(* IEC 61131-3 sources: volt/packages/volt-lsp-iec/test-corpus/pro2193/Device/Plc Logic/Application/09 Misc/Library Manager/L_TB1P_TechnologyBasics, 21 files *)

(* ---- L_TB1P_DIRECTION.dut ---- *)
TYPE L_TB1P_DIRECTION :
(
	DEFAULT := 0,
	CW := 1,
	CCW := 2
);
END_TYPE

(* ---- L_TB1P_STATES.dut ---- *)
TYPE L_TB1P_STATES :
(
	INIT := 1,
	READY := 2,
	CAMMING := 112,
	CAMMING_DONE := 113,
	CLUTCH_OPEN_INSTANT := 114,
	CLUTCH_CLOSE := 115,
	CLUTCH_OPEN := 116,
	CAMSEQUENCER_LOADCAMTABLE := 150,
	CAMSEQUENCER_CYCLICCAM1 := 151,
	CAMSEQUENCER_CYCLICCAM3 := 152,
	CAMSEQUENCER_CAM1CYCLICCAM3CAM1 := 153,
	CAMSEQUENCER_CAM1CAM2CYCLICCAM3CAM4CAM1 := 154,
	ERROR := 999
);
END_TYPE

(* ---- L_TB1P_CONSTANTS.gvl ---- *)
VAR_GLOBAL
	GC_POSITIVE_LIMIT_32BIT : LREAL := 2147483647;
	GC_NEGATIVE_LIMIT_32BIT : LREAL := -2147483647;
END_VAR

(* ---- GETBOOLEANPROPERTY.pou ---- *)
FUNCTION GETBOOLEANPROPERTY : BOOL
VAR_INPUT
	STKEY : WSTRING;
END_VAR
END_FUNCTION

(* ---- GETCOMPANY.pou ---- *)
FUNCTION GETCOMPANY : WSTRING
END_FUNCTION

(* ---- GETNUMBERPROPERTY.pou ---- *)
FUNCTION GETNUMBERPROPERTY : DINT
VAR_INPUT
	STKEY : WSTRING;
END_VAR
END_FUNCTION

(* ---- GETTEXTPROPERTY.pou ---- *)
FUNCTION GETTEXTPROPERTY : WSTRING
VAR_INPUT
	STKEY : WSTRING;
END_VAR
END_FUNCTION

(* ---- GETTEXTPROPERTY2.pou ---- *)
FUNCTION GETTEXTPROPERTY2 : POINTER TO WSTRING
VAR_INPUT
	STKEY : WSTRING;
END_VAR
END_FUNCTION

(* ---- GETTITLE.pou ---- *)
FUNCTION GETTITLE : WSTRING
END_FUNCTION

(* ---- GETVERSION.pou ---- *)
FUNCTION GETVERSION : VERSION
END_FUNCTION

(* ---- GETVERSIONPROPERTY.pou ---- *)
FUNCTION GETVERSIONPROPERTY : VERSION
VAR_INPUT
	STKEY : WSTRING;
END_VAR
END_FUNCTION

(* ---- GLOBALTEXTLIST.pou ---- *)
FUNCTION_BLOCK GLOBALTEXTLIST
VAR
	M_TEXTLISTFILE : STRING(255);
	_STNAMESPACE : STRING;
END_VAR
END_FUNCTION_BLOCK

(* ---- IMAGEPOOL.pou ---- *)
FUNCTION_BLOCK IMAGEPOOL
VAR
	M_STNAMESPACE : STRING(80);
	M_STHELPVARID : STRING;
	M_STHELPVARPATH : STRING(255);
	M_STHELP : STRING;
	M_REGISTERIMAGES : BOOL := TRUE;
END_VAR
END_FUNCTION_BLOCK

METHOD FB_INIT : BOOL
VAR_INPUT
	BINITRETAINS : BOOL;
	BINCOPYCODE : BOOL;
END_VAR
END_METHOD

METHOD FB_REINIT : BOOL
END_METHOD

METHOD FB_EXIT : BOOL
VAR_INPUT
	BINCOPYCODE : BOOL;
END_VAR
END_METHOD

(* ---- L_TB1P_ACCCOMP.pou ---- *)
FUNCTION_BLOCK L_TB1P_ACCCOMP
VAR_INPUT
	LRCYCVEL : LREAL;
	LRMINERTIAMAX : LREAL;
	LRMINERTIACONST : LREAL;
	LRVARIABLEMINERTIA : LREAL;
	LRMINERTIAADAPT : LREAL := 1.0;
	LRFILTERTIMEACCSPEED : REAL := 0.0;
	LRDEADBANDACCTORQUE : LREAL := 0.0;
	LRGAINPOS : LREAL := 1.0;
	LRGAINNEG : LREAL := 1.0;
	XRESET : BOOL;
END_VAR
VAR_OUTPUT
	LRSETACCOUT : LREAL;
	LRSETTORQUEOUT : LREAL;
END_VAR
VAR
	TBDIFFERENTIATE1 : L_USPP_Differentiate;
	LRMINERTIAVAR : LREAL;
	LRLRSETACC_INT : LREAL;
	LRFACTOR_INT : LREAL := 1;
	LRFACTOR : LREAL;
END_VAR
END_FUNCTION_BLOCK

(* ---- L_TB1P_CALCDIAMETER.pou ---- *)
FUNCTION_BLOCK L_TB1P_CALCDIAMETER
VAR_INPUT
	LRCYCREELSPEED : LREAL;
	LRCYCLINEVEL : LREAL;
	LRMAXDIAMETER : LREAL;
	LRMINDIAMETER : LREAL;
	LRCALCULATIONDISTANCE : LREAL := 1;
	XFORCECALCULATION : BOOL;
	XHOLDDIAMETER : BOOL;
	XUNIDIRECT : BOOL;
	XUNWINDACTIVE : BOOL;
	XLOADSETDIAMETER : BOOL;
	LRSETDIAMETER : LREAL;
	LRFILTERTIMEDIAMETER : LREAL := 0;
	LRWINDOWWEBBREAKMONIT : LREAL := 0.1;
END_VAR
VAR_OUTPUT
	XERROR : BOOL;
	EERRORID : L_IE1P_Error;
	LRSETDIAMETEROUT : LREAL;
	LRSETDIAMETERPCTOUT : LREAL;
	LRREZIPRDIAMETERPCT : LREAL;
	XDIAMETERMAXLIMIT : BOOL := FALSE;
	XDIAMETERMINLIMIT : BOOL := FALSE;
	XWEBBREAK : BOOL := FALSE;
	LRMINDIAMETERPCT : LREAL;
	LRSETMINERTIASCALEDOUT : LREAL;
END_VAR
VAR_IN_OUT
	LRDIAMETERRETAIN : LREAL := 0;
END_VAR
VAR
	LRTASKCYCLE : LREAL;
	XTASKCYCLEVALID : BOOL;
	LRFILTERTIME : LREAL;
	LRUNFILTEREDDIAMETER : LREAL;
	LRCALCULATIONDISTANCE_INT : LREAL;
	LRACTSPEEDREEL : LREAL;
	LRNWINDER : LREAL;
	LRREELPOSDIFF : LREAL;
	LRACTPOSDIFF : LREAL;
	LRACTLINESPEED : LREAL;
	LRWICKELWELLENDIFFERENZ : LREAL;
	LRCYCVELLINETMP : LREAL;
	LRSTOREDIAMETER : LREAL;
	LRDIAMETERMONITOR : LREAL;
	LRDIAMETERUNFILTERED : LREAL;
	LRTEMP : LREAL;
	LRTIME : LREAL;
	LRDMAXHYST : LREAL;
	LRDMINHYST : LREAL;
	XRESETCALCINTEGRATORFLAG : BOOL;
	LRMAXDIAMETERINT : LREAL;
	LRMAXDIAMETERMEM : LREAL;
	LRMINDIAMETERINT : LREAL;
	XRETAINLOCAL : BOOL := FALSE;
	LRDIAMETERINT : LREAL;
	LRREFDIAMWEBBREAK : LREAL;
	LRREFDIAMWEBBREAKSCALED : LREAL;
	LRCALCDISTLINEVEL_INT : LREAL;
	LRDIAMETER4CALCDIST : LREAL;
	LRCALCULATIONDISTANCE_OLD : LREAL;
	XHOLDINTEGRATOR_INT : BOOL;
	C_MINDIAMETER : LREAL := 1E-06;
	C_MAXDIAMETER : LREAL := 1000000.0;
	LRLINEVELINTEGRATED : LREAL;
	LRREFDIAMETERWEBBREAK : LREAL;
	LRSETDIAMETERUNFILTERED : LREAL;
	LRWINDERSPEEDINTEGRATED : LREAL;
	XDIAMCALCULATED : BOOL;
	XHOLDINTEGRATOR : BOOL;
END_VAR
END_FUNCTION_BLOCK

METHOD D_MIN_MAX
END_METHOD

METHOD LIMITER
END_METHOD

METHOD SETDIAMETER
VAR_INPUT
	LRNEWDIAMETER : LREAL;
END_VAR
END_METHOD

METHOD FB_INIT : BOOL
VAR_INPUT
	BINITRETAINS : BOOL;
	BINCOPYCODE : BOOL;
END_VAR
END_METHOD

(* ---- L_TB1P_FRICTIONCOMPENSATION.pou ---- *)
FUNCTION_BLOCK L_TB1P_FRICTIONCOMPENSATION
VAR_INPUT
	XIDENT : BOOL;
	XFOLLOWERACTIVE : BOOL;
	LRACTREELSPEEDIN : LREAL;
	LRACTTORQUEIN : LREAL;
	DWSELECTCURVE : DWORD;
	XENABLEFRICTIONCURVE : BOOL;
	LRSETREELSPEED : LREAL;
	LRFRICTIONADAPT : LREAL := 1;
	XINVERTOUTPUT : BOOL;
	LRMAXSPEEDIDENT : LREAL := 10;
	LRACCDECIDENT : LREAL := 1;
	LRFILTERTIMESPEED : LREAL := 0.005;
	LRFILTERTIMETORQUE : LREAL := 0.005;
	LRFILTERTIMEREELSPEED : LREAL := 0.0;
	LRLINEARCOMPSTART : LREAL;
	LRLINEARCOMPEND : LREAL;
	LRLINEARCOMPENDREELSPEED : LREAL;
END_VAR
VAR_OUTPUT
	XBUSY : BOOL;
	XDONE : BOOL;
	XERROR : BOOL := FALSE;
	EERRORID : L_IE1P_Error;
	XSTOP : BOOL;
	XENABLEFOLLOWER : BOOL;
	LRSETREELSPEEDOUT : LREAL;
	LRSETFRICTIONTORQUEOUT : LREAL;
END_VAR
VAR_IN_OUT
	ALRFRICTIONCURVE1 : ARRAY [1..66] OF LREAL;
	ALRFRICTIONCURVE2 : ARRAY [1..66] OF LREAL;
	ALRFRICTIONCURVE3 : ARRAY [1..66] OF LREAL;
	ALRFRICTIONCURVE4 : ARRAY [1..66] OF LREAL;
END_VAR
VAR
	LRTASKCYCLE : LREAL;
	DWINTERNALSTATE : DWORD;
	LRWINDOW : LREAL := 0.001;
	DISTATE : DINT;
	DWFRCURVENO : DWORD;
	XIMPOFF : BOOL;
	XFRICTIONBUSY : BOOL;
	XSTARTFRENABLE : BOOL;
	LRNACTFILTER : LREAL;
	LRMACTFILTER : LREAL;
	LRRAMPVALUE : LREAL;
	LRSTEP : LREAL;
	DWINDEX : DWORD;
	DWNUMBER : DWORD;
	ALRFRICTIONDATA1 : ARRAY [0..64] OF LREAL;
	ALRFRICTIONDATA2 : ARRAY [0..64] OF LREAL;
	LRDIST : LREAL;
	LRHALFDIST : LREAL;
	LRTEMP1 : LREAL;
	LRTEMP2 : LREAL;
	LRNMAXFRICTIONINT : LREAL;
	LRDIFFRAMP : LREAL;
	LRNMAXTIME : LREAL;
	LRACCDECIDENTINT : LREAL;
	LRTIME : LREAL;
	XENABLEFOLLOWEROLD : BOOL;
	LRSPEEDSETFILTER : LREAL;
	LRSPEEDSETFILTERABS : LREAL;
	LRSPEEDSETLIM : LREAL;
	LRDIFFFILTER : LREAL;
	LRACTFRICTION : LREAL;
	LRXTABLEVALUE : LREAL;
	LRMAXVALUE : LREAL;
	LRRESIDUAL : LREAL;
	LRSTRICH : LREAL;
	LRDELTAPOS : LREAL;
END_VAR
END_FUNCTION_BLOCK

METHOD RESETERROR
END_METHOD

(* ---- L_TB1P_IDENTMINERTIA.pou ---- *)
FUNCTION_BLOCK L_TB1P_IDENTMINERTIA
VAR_INPUT
	XIDENT : BOOL;
	XFOLLOWERACTIVE : BOOL;
	LRACTREELSPEEDIN : LREAL;
	LRACTTORQUEIN : LREAL;
	LRMAXSPEEDIDENT : LREAL := 10;
	LRMAXTORQUEIDENT : LREAL := 1;
	LRFILTERTIMESPEED : LREAL := 0.005;
	LRFILTERTIMETORQUE : LREAL := 0.005;
	LRFILTERTIMEREELSPEED : LREAL := 0.0;
END_VAR
VAR_OUTPUT
	XBUSY : BOOL;
	XDONE : BOOL;
	XERROR : BOOL := FALSE;
	EERRORID : L_IE1P_Error;
	XENABLEFOLLOWER : BOOL;
	LRSETTORQUEOUT : LREAL;
	LRMINERTIAIDENT : LREAL;
END_VAR
VAR
	LRMINERTIAMAXTOLERANCEERROR : LREAL;
	LRTASKCYCLE : LREAL;
	DWINTERNALSTATE : DWORD;
	DWINDEX : DWORD;
	DISTATE : DINT;
	XIMPOFF : BOOL;
	XACTIVE : BOOL;
	XMINERTIABUSY : BOOL;
	LRNACTFILTER : LREAL;
	LRMACTFILTER : LREAL;
	LRTIME : LREAL;
	LRNMAXMOTORINTERN : LREAL;
	LRMMAXMOTORINTERN : LREAL;
	LRNACTAKKU : LREAL;
	LRMACTAKKU : LREAL;
	LRSIGNNMAX : LREAL := 1;
	LRMSETMINERTIAINT_N : LREAL;
	LRNMAXMINERTIAINT_N : LREAL;
	LRACCTIME : LREAL;
	LRDECTIME : LREAL;
	LRTOTALTIME : LREAL;
	LRWAITTIME : LREAL;
END_VAR
END_FUNCTION_BLOCK

METHOD RESETERROR
END_METHOD

(* ---- L_TB1P_MARKREGISTER.pou ---- *)
FUNCTION_BLOCK L_TB1P_MARKREGISTER
VAR_INPUT
	XENABLE : BOOL;
	LRCYCSETVEL : LREAL;
	XTPRECEIVEDIN : BOOL;
	LRSETTPDIFFERENCE : LREAL;
	LRMARKSTACKLENGTH : LREAL;
	XCORRECTIONBUSY : BOOL;
	LRSETPOSCORRIN : LREAL;
END_VAR
VAR_OUTPUT
	XTPRECEIVEDOUT : BOOL;
	LRTPDIFFERENCEOUT : LREAL;
	LRTOTALSTACKDIFFERENCEOUT : LREAL;
	XERROR : BOOL := FALSE;
	EERRORID : L_IE1P_Error;
END_VAR
VAR
	LRTPDIFFERENCES : ARRAY [1..64] OF LREAL := [64(0)];
	LRTPPOSITION : ARRAY [1..64] OF LREAL := [64(0)];
	XTPVALID : ARRAY [1..64] OF BOOL := [64(FALSE)];
	SDINTEGRATEAXIS1 : L_MC1P_IntegrateAxis;
	COUNTERIN : WORD := 1;
	COUNTEROUT : WORD := 1;
	DWINTEGRATORVALUE : DWORD := 0;
	LRINTEGRATORPOS : LREAL := 0;
	LRTASKCYCLE : LREAL;
	LRPOSDIFF : LREAL;
	LRPOSTOREGISTEREND : LREAL;
	XREGISTERFULL : BOOL;
	LRPOSDIFFINSTACK : LREAL := 0;
	DWCOUNTER : DWORD;
	XINIT : BOOL;
	XWAITINGFORCORRECTIONDONE : BOOL;
	XCORRETIONSTARTED : BOOL;
	LRACTUALTPDIFFERENCE : LREAL;
	XCORRECTIONBUSY_OLD : BOOL;
	LRSETPOSCORRIN_OLD : LREAL;
END_VAR
END_FUNCTION_BLOCK

METHOD CALL_CALCULATETOTALSTACK
END_METHOD

METHOD CALL_WAITFORCORRECTION
END_METHOD

(* ---- L_TB1P_MARKWINDOW.pou ---- *)
FUNCTION_BLOCK L_TB1P_MARKWINDOW
VAR_INPUT
	XENABLE : BOOL;
	LRCYCREGISTERPOS : LREAL;
	LRCYCSETVEL : LREAL;
	XTPRECEIVEDIN : BOOL;
	LRACTTPPOSIN : LREAL;
	XTEACHMARKWINDOW : BOOL;
	LRSETMARKDISTANCE : LREAL;
	LRMARKSENSORPOSITION : LREAL;
	LRSETMARKWINDOW : LREAL;
	LRSETOFFSETMARKWINDOW : LREAL;
	DWMAXTPNOTDETECTED : DWORD;
END_VAR
VAR_OUTPUT
	XTPRECEIVEDOUT : BOOL;
	XTPWINDOWOPEN : BOOL;
	XTPWINDOWOPENCOMP : BOOL;
	LRTPDELTAPOSCOMP : LREAL;
	XTPINWINDOW : BOOL;
	XTPNOTINWINDOW : BOOL;
	XTPNOTDETECTED : BOOL;
	XTPSENSORTEACHED : BOOL;
	LRACTTPPOS : LREAL;
	XMAXTPNOTDETECTED : BOOL;
END_VAR
VAR
	XFIRSTSENSOR : BOOL;
	XTPWINDOWOPENOLD : BOOL;
	XTPNOTDETECTEDINTERNAL : BOOL;
	LRLOWERWINDOW : LREAL;
	LRUPPERWINDOW : LREAL;
	LRTPPOSINWINDOWTEST : LREAL;
	XTEACHTPSENSOROLD : BOOL;
	DWMISSEDTPCOUNTER : DWORD;
	LRACTUALREGISTERPOS : LREAL;
	XTPISINWINDOW : BOOL;
	XMISSEDTPDECREMENT : BOOL;
	LRDEADTIMEPOSDIFF : LREAL;
	LRUPPERWINDOWCOMP : LREAL;
	XTPCOMPWINDOWOPEN : BOOL;
	XTPCOMPWINDOWOPENOLD : BOOL := FALSE;
	LRLOWERWINDOWCOMP : LREAL;
	XTPRECEIVEDOLD : BOOL;
	LRACTUALREGISTERPOSOLD : LREAL;
	XTPRECEIVEDINTERNAL : BOOL;
	LRTASKCYCLE : LREAL;
END_VAR
END_FUNCTION_BLOCK

(* ---- L_TB1P_POSDIFFCORRECTION.pou ---- *)
FUNCTION_BLOCK L_TB1P_POSDIFFCORRECTION
VAR_INPUT
	XENABLE : BOOL;
	LRCYCSETVEL : LREAL;
	XLOADSTARTPOS : BOOL;
	LRSTARTPOS : LREAL;
	XTPRECEIVEDIN : BOOL;
	LRSETCORRECTION : LREAL;
	XCORRWINDOWINXUNITS : BOOL;
	LRSETUPPERWINDOW : LREAL;
	LRSETLOWERWINDOW : LREAL;
	LRCYCPOSFEEDBACK : LREAL;
	DNSETNUMERATORAXISY : DWORD := 1;
	DNSETDENOMINATORAXISY : DWORD := 1;
	LRSETCYCLELENGTHX : LREAL;
	LRSETCYCLELENGTHY : LREAL;
END_VAR
VAR_OUTPUT
	XBUSY : BOOL;
	XCORRECTIONBUSY : BOOL;
	LRSETPOSOUT : LREAL;
	LRSETINTEGRATEDPOSITION : LREAL;
	LRSETPOSCORROUT : LREAL;
	XERROR : BOOL;
	EERRORID : L_IE1P_Error;
END_VAR
VAR_IN_OUT
	AXIS : AXIS_REF;
END_VAR
VAR
	LRDELTAPOSTOTAL : LREAL;
	LRMASTERDISTANCE : LREAL;
	LRPOSITIONSET : LREAL;
	LRPOSITIONNORMED : LREAL;
	LRPOSITIONOUTNORMED : LREAL;
	LRDELTAPOSCORRECTION : LREAL;
	LRPOSITIONSETOLD : LREAL;
	LRPOSITIONSETAXISOUT : LREAL;
	BYSTEPPER : BYTE;
	LRCORRECTIONDISTANCELOCAL : LREAL;
	LRCORRECTIONLOCAL : LREAL;
	L_DIFFERENTIATE : L_MC2P_Differentiate;
	INTEGRATOR : L_MC1P_IntegrateAxis;
	LRDELTAPOSOUT : LREAL;
	XEXECUTECORRECTIONINTERN : BOOL;
	XPOSITIVEDIRECTION : BOOL := FALSE;
	LRCORRECTIONDISTANCE : LREAL;
	LRUPPERWINDOWINTERNAL : LREAL;
	LRLOWERWINDOWINTERNAL : LREAL;
	FTASKCYCLE : LREAL;
	XCORRECTIONACTIVE : BOOL;
	LRCORRECTIONLOCAL1 : LREAL;
	XTPRECEIVEDOLD : BOOL;
	LRINTEGRATORSPEED : LREAL;
	XWINDOWINCYCLE : BOOL;
	LRDELTAWINDOW : LREAL;
	LRCYCPOSINTOOLINTERNAL : LREAL;
	LRUPPERWINDOWINTERNALDELTA : LREAL;
	LRLOWERWINDOWINTERNALDELTA : LREAL;
	XINIT : BOOL := TRUE;
	XINITOUTOFCORRWINDOW : BOOL := TRUE;
	LRLOWERWINDOWINTERNALOLD : LREAL;
	LRUPPERWINDOWINTERNALOLD : LREAL;
	LRCYCPOSFEEDBACKINT : LREAL;
	XCORRECTIONBUSYOLD : BOOL;
	LRSETPOSCORROUTOLD : LREAL;
	LRCYCPOSINTOOLINTERNAL_CASE : LREAL;
	XWINDOWCHANGEDFLAG : BOOL := FALSE;
END_VAR
END_FUNCTION_BLOCK

(* ---- L_TB1P_TENSIONCURVE.pou ---- *)
FUNCTION_BLOCK L_TB1P_TENSIONCURVE
VAR_INPUT
	XENABLE : BOOL;
	LRSETTENSIONIN : LREAL;
	DWSELECTCURVE : DWORD;
	LRCURVECTRLSCALED : LREAL;
	LRSTARTDIAMETERPCT : LREAL;
	LRSETDIAMETERPCT : LREAL;
	ALRTENSIONCURVE : ARRAY [1..65] OF LREAL;
END_VAR
VAR_OUTPUT
	LRSETTENSIONOUT : LREAL;
	LRCURVEVALUESCALED : LREAL;
END_VAR
VAR
	LRTEMP : LREAL;
	LRTEMP1 : LREAL;
	LRTEMP2 : LREAL;
	LRXTABLEVALUE : LREAL;
	DWINDEX : DWORD;
	LRRESIDUAL : LREAL;
	DWSELECTCURVE_INT : DWORD;
	LRDIAMETER_INT : LREAL;
	LRCURVECTRL_INT : LREAL;
	LRSTARTDIAMETER_INT : LREAL;
	LRSTRICH : LREAL;
	LRDELTAPOS : LREAL;
END_VAR
END_FUNCTION_BLOCK
